(* IEC 61131-3 sources: 2026_Projet_YGO_ExcavatriceDragage/CODE_BACKUP/CODE_20260807_v0.5.25/COMMUN, 15 files *)

(* ---- E_State.st ---- *)
(* ═══════════════════════════════════════════════════════════════
   🚦 E_State — Phase opérationnelle d'un FB métier (valeurs EXCLUSIVES)
   ───────────────────────────────────────────────────────────────
    📄 Doc métier : DOC/AF_Partie-03_Contrats_Composants_v2.1.md §3
   ⚠️ Un seul état à la fois. Error / SafeStop / perte Enable sont
      ORTHOGONAUX à la phase (voir ErrorId, ne polluent pas State).
   🧩 Fondation manquante requise par le contrat FB (Partie3 §1).
   ═══════════════════════════════════════════════════════════════ *)

TYPE E_State :
ENUM
    DISABLED := 0,   (* Enable faux, neutralisé *)
    INIT     := 1,   (* Démarrage / vérifs *)
    READY    := 2,   (* Prêt, attend ordre *)
    BUSY     := 3,   (* Action en cours *)
    DONE     := 4,   (* Action terminée *)
    STOPPING := 5    (* Décél rampe avant arrêt (StartStop=FALSE ou SafeStop=TRUE) *)
END_ENUM
END_TYPE

(* ---- ST_ContactorCheck.st ---- *)
(* ═══════════════════════════════════════════════════════════════
   🔌 ST_ContactorCheck — Double vérification commande/retour contacteur
   ───────────────────────────────────────────────────────────────
    📄 Doc métier : DOC/AF_Partie-02_Architecture_Programme_v3.1.md §3,
                    DOC/AF_Partie-03_Contrats_Composants_v2.1.md §2
   Utilisé par FB_Brake (frein) et FB_Winch (contacteurs de sens) pour
   détecter un collage / une absence de fermeture d'un contacteur de
   puissance, au-delà d'un délai de cohérence (FeedbackTimeout du FB
   appelant).
   ═══════════════════════════════════════════════════════════════ *)

TYPE ST_ContactorCheck :
STRUCT
    Command     : BOOL;   // Ordre envoyé au contacteur (TRUE = fermé/actif)
    Feedback    : BOOL;   // Retour d'état câblé (TRUE = effectivement fermé)
    StuckClosed : BOOL;   // Diag : commande OFF mais retour ON depuis trop longtemps → PowerCutOff
    StuckOpen   : BOOL;   // Diag : commande ON mais retour OFF depuis trop longtemps
END_STRUCT
END_TYPE

(* ---- FB_Acquisition_Preflight.st ---- *)
(* ═══════════════════════════════════════════════════════════════
   🩺 FB_Acquisition_Preflight — Verdict passif machine arrêtée
   📄 Doc : ARCHIVES/Doc/AUDITS/PreLivraison/TASKS/TASK_D1_Preflight_et_Symetrie_Winch_v1.0.md
   🔒 Observateur pur : aucun SafeStop, PowerCutOff ou ordre machine.
   ═══════════════════════════════════════════════════════════════ *)
FUNCTION_BLOCK FB_Acquisition_Preflight
VAR_INPUT
    Execute : BOOL;
    MachineIsStill : BOOL;
    M1BrakeApplied, M2BrakeApplied, M3BrakeApplied : BOOL;
    M1ContactorsReleased, M2ContactorsReleased, M1ThermalOk, M2ThermalOk : BOOL;
    BrakeThermalOk, PhaseRotationOk, SlackCableTensioned, M3SensorWordIncoherent : BOOL;
    EmergencyChainClosed, PowerContactorEngaged, EncoderM1Operational, EncoderM2Operational : BOOL;
    HomedM1, HomedM2, M1PositionInBounds, M2PositionInBounds : BOOL;
END_VAR
VAR_OUTPUT
    PreflightOk : BOOL;
    PreflightDone : BOOL;
    PreflightBusy : BOOL;
    PreflightErrorId : WORD;
END_VAR
VAR
    ExecuteEdge : R_TRIG;
    BootPending : BOOL := TRUE;
    RequestPending : BOOL;
END_VAR

ExecuteEdge(CLK := Execute);
RequestPending := RequestPending OR ExecuteEdge.Q OR BootPending;
PreflightBusy := RequestPending AND NOT MachineIsStill;
IF NOT MachineIsStill THEN PreflightDone := FALSE; RETURN; END_IF;
IF NOT RequestPending THEN RETURN; END_IF;

PreflightErrorId := 0;
(* bit0..2 frein M1/M2/M3 serré; bit3..4 contacteurs M1/M2 retombés;
   bit5..6 thermique M1/M2 OK; bit7 thermique frein OK; bit8 phases OK;
   bit9 câble M2 tendu; bit10 mot M3 cohérent; bit11 contacteur sans chaîne;
   bit12..13 codeur M1/M2 opérationnel; bit14..15 homé et position bornée M1/M2. *)
IF NOT M1BrakeApplied THEN PreflightErrorId := PreflightErrorId OR 16#0001; END_IF;
IF NOT M2BrakeApplied THEN PreflightErrorId := PreflightErrorId OR 16#0002; END_IF;
IF NOT M3BrakeApplied THEN PreflightErrorId := PreflightErrorId OR 16#0004; END_IF;
IF NOT M1ContactorsReleased THEN PreflightErrorId := PreflightErrorId OR 16#0008; END_IF;
IF NOT M2ContactorsReleased THEN PreflightErrorId := PreflightErrorId OR 16#0010; END_IF;
IF NOT M1ThermalOk THEN PreflightErrorId := PreflightErrorId OR 16#0020; END_IF;
IF NOT M2ThermalOk THEN PreflightErrorId := PreflightErrorId OR 16#0040; END_IF;
IF NOT BrakeThermalOk THEN PreflightErrorId := PreflightErrorId OR 16#0080; END_IF;
IF NOT PhaseRotationOk THEN PreflightErrorId := PreflightErrorId OR 16#0100; END_IF;
IF NOT SlackCableTensioned THEN PreflightErrorId := PreflightErrorId OR 16#0200; END_IF;
IF M3SensorWordIncoherent THEN PreflightErrorId := PreflightErrorId OR 16#0400; END_IF;
IF PowerContactorEngaged AND NOT EmergencyChainClosed THEN PreflightErrorId := PreflightErrorId OR 16#0800; END_IF;
IF NOT EncoderM1Operational THEN PreflightErrorId := PreflightErrorId OR 16#1000; END_IF;
IF NOT EncoderM2Operational THEN PreflightErrorId := PreflightErrorId OR 16#2000; END_IF;
IF NOT HomedM1 OR NOT M1PositionInBounds THEN PreflightErrorId := PreflightErrorId OR 16#4000; END_IF;
IF NOT HomedM2 OR NOT M2PositionInBounds THEN PreflightErrorId := PreflightErrorId OR 16#8000; END_IF;
PreflightOk := (PreflightErrorId = 0); PreflightDone := TRUE; BootPending := FALSE; RequestPending := FALSE;

(* ---- FB_Brake.st ---- *)
(* ═══════════════════════════════════════════════════════════════
   🛑 FB_Brake — Séquence frein à manque de courant (temps physiques)
   ───────────────────────────────────────────────────────────────
   📄 Doc métier : DOC/AF_Partie-10_Fonction_Winch_v2.0.md §3
                   (règles issues de DOC/AF_Partie-04_Mode_SemiAuto_Sequenceur_v2.0.md §4)
   🛠️ Frein à manque de courant : colle au repos (sécurité positive).
   📥 MovementRequested : mouvement demandé par FB_Winch (sens+palier > 0)
   📤 BrakeCmd          : commande bobine frein — TRUE = relâché (alimenté)
   ⏱️ Séquence démarrage : attend fermeture contacteur + magnétisation
      moteur AVANT de relâcher (sinon charge retombe → à-coup).
   ⏱️ Séquence arrêt     : attend décélération/ouverture contacteur AVANT
      de coller (sinon usure/casse mécanique en plein mouvement).
   🔍 Double vérification retour contacteur bobine (ST_ContactorCheck) :
      incohérence commande/retour au-delà de FeedbackTimeout → ErrorId.
   🆕 REX 2026-08-03 (révocation 2026-07-26) : le retour câblé est l'image du CONTACTEUR DE COMMANDE
      (DI = 1 ⟺ frein ouvert). Plus d'inversion à la frontière : ce FB reçoit maintenant un
      signal dans le MÊME sens que `BrakeCmd` en marche saine (TRUE = relâché = ouvert) → le test d'incohérence est `<>`, pas `=`.
      ⚠️ Ce retour n'est PAS une mesure du frein : il détecte un contacteur/bobine défaillant, mais
      pas un frein usé ou qui patine. Le patinage reste couvert par Méca A (dérive codeur,
      FB_Safety_Winch bit7) — pas par ce bloc.
   ═══════════════════════════════════════════════════════════════ *)

// === DECLARATION (à coller dans la partie déclaration du POU FB_Brake) ===

FUNCTION_BLOCK PUBLIC FB_Brake
VAR_INPUT
    Enable              : BOOL;                     // Contexte général (comme tout FB) — FALSE = frein collé (sûr)
    Reset               : BOOL;                     // Acquittement défaut (front)
    MovementRequested   : BOOL;                      // TRUE = FB_Winch demande un mouvement (sens+palier actifs)
    ContactorFeedback   : BOOL;                      // Retour frein (`PRG_02_Acquisition.HwIn`) : TRUE = frein OUVERT (desserré)
                                                       // 🆕 REX 2026-08-03 : même sens que BrakeCmd (TRUE = relâché)
                                                       // → en marche normale les deux sont ÉGAUX ; c'est leur
                                                       //   DIFFÉRENCE qui trahit un contacteur collé (voir §4).
    DelayContactClose   : TIME := T#100ms;            // Temps de fermeture contacteur de puissance
    DelayMagnetise      : TIME := T#300ms;            // Délai magnétisation moteur avant ouverture frein
    DelayMotorDecel     : TIME := T#500ms;            // Délai décélération/ouverture contacteur avant collage frein
    FeedbackTimeout     : TIME := T#1s;               // Délai max cohérence commande/retour frein
    BypassContactorCheck: BOOL;                       // 🧪 TRUE = désactive StuckClosed/StuckOpen (axe simulé,
                                                       // voir GVL_Simulation.SensorMxContactorFeedbackIsReal, passé
                                                       // par l'appelant FB_Winch/FB_Translation — TOUJOURS FALSE réel)
END_VAR
VAR_OUTPUT
    Ready               : BOOL;
    Busy                : BOOL;
    Done                : BOOL;
    Error               : BOOL;
    ErrorId             : WORD;          // bit0: "Défaut engagement frein" - incohérence commande/retour frein (collage ou non-relâche)
    State               : E_State;
    StateAtError        : E_State;
    BrakeCmd            : BOOL;          // Commande sortie bobine frein : TRUE = relâché
    BrakeCommandOpenConfirmed : BOOL;    // TRUE = frein ouvert = commande ouverture confirmée (même sens que ContactorFeedback)
    ContactorCheck      : ST_ContactorCheck;  // Diag détaillé (IHM / FB_Safety_Winch)
END_VAR
VAR
    ResetEdge           : R_TRIG;
    ErrorEdge           : R_TRIG;
    BypassEdge          : R_TRIG;        // 🔑 REX 2026-07-24 : Front montant activation bypass pour réarmement immédiat
    TonMagnetise        : TON;           // Temporisation avant relâche
    TonDecel            : TON;           // Temporisation avant collage
    TonFeedback         : TON;           // Timeout cohérence commande/retour
END_VAR

// === IMPLEMENTATION (à coller dans le corps ST du POU FB_Brake) ===

// 🛑 1. GATE — pas d'Enable = frein collé (sécurité positive), aucune temporisation en cours
IF NOT Enable THEN
    TonMagnetise(IN := FALSE, PT := DelayMagnetise + DelayContactClose);
    TonDecel(IN := FALSE, PT := DelayMotorDecel);
    BrakeCmd := FALSE;
    State := E_State.DISABLED;
    Ready := FALSE; Busy := FALSE; Done := FALSE;
    RETURN;
END_IF;

Ready := TRUE;

// 🔑 2. RESET FRONT — efface le bit dont la cause a disparu
ResetEdge(CLK := Reset);
BypassEdge(CLK := BypassContactorCheck);

// 🛠️ 3. SÉQUENCE TEMPORISÉE (démarrage vs arrêt)
IF MovementRequested THEN
    TonDecel(IN := FALSE, PT := DelayMotorDecel);
    TonMagnetise(IN := TRUE, PT := DelayMagnetise + DelayContactClose);
    IF TonMagnetise.Q THEN
        BrakeCmd := TRUE;              // ✅ Contacteur + magnétisation acquis → relâche
        State := E_State.DONE;
    ELSE
        BrakeCmd := FALSE;             // ⏳ Encore collé pendant la magnétisation
        State := E_State.BUSY;
    END_IF;
ELSE
    // 🆕 REX 2026-07-08 : Sécurité positive - fermeture immédiate du frein (collé) dès que les contacteurs de sens s'ouvrent
    TonMagnetise(IN := FALSE, PT := DelayMagnetise + DelayContactClose);
    TonDecel(IN := FALSE, PT := DelayMotorDecel);
    BrakeCmd := FALSE;                 // Fermeture immédiate
    State := E_State.READY;
END_IF;

Busy := (State = E_State.BUSY);
Done := (State = E_State.DONE);

// 🔍 4. DOUBLE VÉRIFICATION RETOUR CONTACTEUR (ST_ContactorCheck)
ContactorCheck.Command := BrakeCmd;
ContactorCheck.Feedback := ContactorFeedback;

// 🆕 REX 2026-08-03 (révocation 2026-07-26) : `ContactorFeedback` est maintenant dans le MÊME sens
// que `BrakeCmd` (TRUE = relâché = frein ouvert). En marche saine les deux sont ÉGAUX → c'est leur
// DIFFÉRENCE qui signale l'incohérence (contacteur collé).
// ⚠️ Le test repasse en `<>` (retour à la logique d'origine pré-2026-07-26).
TonFeedback(IN := (BrakeCmd <> ContactorFeedback), PT := FeedbackTimeout);
IF NOT BypassContactorCheck THEN
    IF TonFeedback.Q THEN
        ContactorCheck.StuckClosed := (BrakeCmd AND NOT ContactorFeedback);            // relâche commandée (BrakeCmd=TRUE), frein reste serré (ContactorFeedback=FALSE)
        ContactorCheck.StuckOpen   := (NOT BrakeCmd AND ContactorFeedback);             // serrage commandé (BrakeCmd=FALSE), frein reste ouvert (ContactorFeedback=TRUE)
        ErrorId := ErrorId OR 16#0001;
    ELSIF ResetEdge.Q THEN
        ContactorCheck.StuckClosed := FALSE;
        ContactorCheck.StuckOpen   := FALSE;
        ErrorId := ErrorId AND 16#FFFE;
    END_IF;
ELSE
    ContactorCheck.StuckClosed := FALSE;
    ContactorCheck.StuckOpen   := FALSE;
    ErrorId := ErrorId AND 16#FFFE;   // Bypass actif : efface/maintient à 0 le bit 0
    IF BypassEdge.Q THEN
        StateAtError := E_State.DISABLED; // Front activation bypass : débloque l'état figé
    END_IF;
END_IF;

// 🧾 5. ARBITRAGE ERROR / STATEATERROR (figé jusqu'à acquittement)
Error := (ErrorId <> 16#0000);
ErrorEdge(CLK := Error);
IF ErrorEdge.Q THEN
    StateAtError := State;
END_IF;

// 🛡️ 6. SORTIE SÛRE SUR DÉFAUT
IF Error THEN
    BrakeCmd := FALSE;
END_IF;

// 📤 7. CONFIRMATION OUVERTURE FREIN (même sens que ContactorFeedback, ou image de BrakeCmd si BypassContactorCheck=TRUE)
IF BypassContactorCheck THEN
    BrakeCommandOpenConfirmed := BrakeCmd;
ELSE
    BrakeCommandOpenConfirmed := ContactorFeedback;  (* TRUE = frein ouvert = desserrage confirmé *)
END_IF;

(* ---- FB_CfgPersistBridge_BucketCfg.st ---- *)
(* ═══════════════════════════════════════════════════════════════
   🌉 FB_CfgPersistBridge_BucketCfg — Pont persistance générique pour ST_BucketCfg
   ───────────────────────────────────────────────────────────────
   🎯 Voir FB_CfgPersistBridge_SyncCfg.st (Lot 3a) pour la logique de référence — identique,
   seul le type ST_BucketCfg change. La copie struct-à-struct gère aussi le sous-struct imbriqué
   Config : ST_BucketConfig automatiquement (pas de traitement spécial nécessaire).
   ═══════════════════════════════════════════════════════════════ *)
FUNCTION_BLOCK FB_CfgPersistBridge_BucketCfg
VAR_IN_OUT
    Hmi     : ST_BucketCfg; (* 🖥️ ex. GVL_IHM.M2TreuilBenne.Bucket.Cfg *)
    Persist : ST_BucketCfg; (* 💾 ex. GVL_PERSISTENT._BucketCfgPersist *)
END_VAR
VAR_OUTPUT
    JustRestored : BOOL;
END_VAR

JustRestored := FALSE;
IF NOT Hmi.Initialized THEN
    Hmi := Persist;
    Hmi.Initialized := TRUE;
    JustRestored := TRUE;
ELSE
    Persist := Hmi;
END_IF;

(* ---- FB_CfgPersistBridge_CommunCfg.st ---- *)
(* ═══════════════════════════════════════════════════════════════
   🌉 FB_CfgPersistBridge_CommunCfg — Pont persistance générique pour ST_CommunCfg
   ───────────────────────────────────────────────────────────────
   🎯 Voir FB_CfgPersistBridge_SyncCfg.st (Lot 3a) pour la logique de référence — identique,
   seul le type ST_CommunCfg change.
   ═══════════════════════════════════════════════════════════════ *)
FUNCTION_BLOCK FB_CfgPersistBridge_CommunCfg
VAR_IN_OUT
    Hmi     : ST_CommunCfg; (* 🖥️ ex. GVL_IHM.Commun.Cfg *)
    Persist : ST_CommunCfg; (* 💾 ex. GVL_PERSISTENT._CommunCfgPersist *)
END_VAR
VAR_OUTPUT
    JustRestored : BOOL;
END_VAR

JustRestored := FALSE;
IF NOT Hmi.Initialized THEN
    Hmi := Persist;
    Hmi.Initialized := TRUE;
    JustRestored := TRUE;
ELSE
    Persist := Hmi;
END_IF;

(* ---- FB_CfgPersistBridge_CycleCfg.st ---- *)
(* ═══════════════════════════════════════════════════════════════
   🌉 FB_CfgPersistBridge_CycleCfg — Pont persistance générique pour ST_CycleCfg
   ───────────────────────────────────────────────────────────────
   🎯 Voir FB_CfgPersistBridge_SyncCfg.st (Lot 3a) pour la logique de référence — identique,
   seul le type ST_CycleCfg change.
   ═══════════════════════════════════════════════════════════════ *)
FUNCTION_BLOCK FB_CfgPersistBridge_CycleCfg
VAR_IN_OUT
    Hmi     : ST_CycleCfg; (* 🖥️ ex. GVL_IHM.Cycle.Cfg *)
    Persist : ST_CycleCfg; (* 💾 ex. GVL_PERSISTENT._CycleCfgPersist *)
END_VAR
VAR_OUTPUT
    JustRestored : BOOL;
END_VAR

JustRestored := FALSE;
IF NOT Hmi.Initialized THEN
    Hmi := Persist;
    Hmi.Initialized := TRUE;
    JustRestored := TRUE;
ELSE
    Persist := Hmi;
END_IF;

(* ---- FB_CfgPersistBridge_DredgingAssistCfg.st ---- *)
(* ═══════════════════════════════════════════════════════════════
   🌉 FB_CfgPersistBridge_DredgingAssistCfg — Pont IHM/persistance prélèvement
   ═══════════════════════════════════════════════════════════════ *)
FUNCTION_BLOCK FB_CfgPersistBridge_DredgingAssistCfg
VAR_IN_OUT
    Hmi     : ST_DredgingAssistCfg;
    Persist : ST_DredgingAssistCfg;
END_VAR
VAR_OUTPUT
    JustRestored : BOOL;
END_VAR

JustRestored := FALSE;
IF NOT Hmi.Initialized THEN
    Hmi := Persist;
    Hmi.Initialized := TRUE;
    JustRestored := TRUE;
ELSE
    Persist := Hmi;
END_IF;

(* ---- FB_CfgPersistBridge_SyncCfg.st ---- *)
(* ═══════════════════════════════════════════════════════════════
   🌉 FB_CfgPersistBridge_SyncCfg — Pont persistance générique pour ST_SyncCfg
   ───────────────────────────────────────────────────────────────
   🎯 Remplace les blocs manuels restauration/sauvegarde dupliqués à chaque domaine
   (voir DOC/AUDITS/ConfigPersistence/). Une instance = un couple (struct IHM, struct
   GVL_PERSISTENT) du MÊME type. Logique :
   - Hmi.Initialized = FALSE (RETAIN invalidé, ex. changement de layout DUT) → restaure
     Hmi depuis Persist, marque Initialized, pulse JustRestored 1 scan.
   - Hmi.Initialized = TRUE → sauvegarde continue Hmi vers Persist (jamais l'inverse).
   🔒 Défense en profondeur : jamais d'écriture PERSISTENT avant qu'une restauration
   réussie n'ait eu lieu (même principe que tous les blocs Cfg du Lot 2).
   ═══════════════════════════════════════════════════════════════ *)
FUNCTION_BLOCK FB_CfgPersistBridge_SyncCfg
VAR_IN_OUT
    Hmi     : ST_SyncCfg; (* 🖥️ ex. GVL_IHM.M1M2Sync.Cfg — struct exposé à l'IHM *)
    Persist : ST_SyncCfg; (* 💾 ex. GVL_PERSISTENT._SyncCfgPersist — mémoire PERSISTENT *)
END_VAR
VAR_OUTPUT
    JustRestored : BOOL; (* 🔔 TRUE pendant 1 scan le boot où la restauration a eu lieu —
                             l'appelant s'en sert pour piloter GVL_IHM.Commun.ConfigRestoredFromPersistent *)
END_VAR

JustRestored := FALSE;
IF NOT Hmi.Initialized THEN
    Hmi := Persist;
    Hmi.Initialized := TRUE;
    JustRestored := TRUE;
ELSE
    Persist := Hmi;
END_IF;

(* ---- FB_CfgPersistBridge_TranslationCfg.st ---- *)
(* ═══════════════════════════════════════════════════════════════
   🌉 FB_CfgPersistBridge_TranslationCfg — Pont persistance générique pour ST_TranslationCfg
   ───────────────────────────────────────────────────────────────
   🎯 Instance unique : TranslationM3.Cfg (un seul axe M3, contrairement à M1/M2).
   Restaure Persist → Hmi au boot si nécessaire, puis sauvegarde Hmi → Persist.
   ═══════════════════════════════════════════════════════════════ *)
FUNCTION_BLOCK FB_CfgPersistBridge_TranslationCfg
VAR_IN_OUT
    Hmi     : ST_TranslationCfg; (* 🖥️ Struct exposé à l'IHM *)
    Persist : ST_TranslationCfg; (* 💾 Mémoire PERSISTENT *)
END_VAR
VAR_OUTPUT
    JustRestored : BOOL; (* 🔔 TRUE pendant le scan de restauration *)
END_VAR

JustRestored := FALSE;
IF NOT Hmi.Initialized THEN
    Hmi := Persist;
    Hmi.Initialized := TRUE;
    JustRestored := TRUE;
ELSE
    Persist := Hmi;
END_IF;

(* ---- FB_CfgPersistBridge_WinchCfg.st ---- *)
(* ═══════════════════════════════════════════════════════════════
   🌉 FB_CfgPersistBridge_WinchCfg — Pont persistance générique pour ST_WinchCfg
   ───────────────────────────────────────────────────────────────
   🎯 Deux instances indépendantes : M1TreuilRetenue.Cfg et M2TreuilBenne.Cfg.
   Restaure Persist → Hmi au boot si nécessaire, puis sauvegarde Hmi → Persist.
   ═══════════════════════════════════════════════════════════════ *)
FUNCTION_BLOCK FB_CfgPersistBridge_WinchCfg
VAR_IN_OUT
    Hmi     : ST_WinchCfg; (* 🖥️ Struct exposé à l'IHM *)
    Persist : ST_WinchCfg; (* 💾 Mémoire PERSISTENT *)
END_VAR
VAR_OUTPUT
    JustRestored : BOOL; (* 🔔 TRUE pendant le scan de restauration *)
END_VAR

JustRestored := FALSE;
IF NOT Hmi.Initialized THEN
    Hmi := Persist;
    Hmi.Initialized := TRUE;
    JustRestored := TRUE;
ELSE
    Persist := Hmi;
END_IF;

(* ---- FB_CycleTime.st ---- *)
(* ═══════════════════════════════════════════════════════════════
   ⏱️ FB_CycleTime — Mesure du temps de cycle réel de la tâche
   ───────────────────────────────────────────────────────────────
   📄 Doc métier : DOC/AF_Partie-08_Fonction_Joystick_v2.0.md §2
      (base de temps utilisée par FB_Filter_PT1, composé dans FB_Joystick)
   ═══════════════════════════════════════════════════════════════ *)
FUNCTION_BLOCK FB_CycleTime
VAR_INPUT
    DefaultValueS : REAL := 0.004; (* Valeur de secours par défaut (ex. 4ms) *)
END_VAR
VAR_OUTPUT
    CycleTimeS    : REAL;          (* Temps écoulé réel calculé (secondes) *)
END_VAR
VAR
    TimeCurrent   : TIME;          (* Temps système actuel *)
    TimeLast      : TIME;          (* Empreinte de temps du cycle précédent *)
    DeltaTimeMs   : UDINT;         (* Écart brut calculé (ms) *)
    InitDone      : BOOL;          (* Drapeau d'initialisation du premier cycle *)
END_VAR

// 1. ACQUISITION DU TEMPS SYSTÈME
TimeCurrent := TIME();

// 2. INITIALISATION UNIQUE AU PREMIER CYCLE
IF NOT InitDone THEN
    TimeLast := TimeCurrent;
    InitDone := TRUE;
    CycleTimeS := DefaultValueS;
    RETURN;
END_IF;

// 3. CALCUL DU DELTA EN MILLISECONDES
DeltaTimeMs := TIME_TO_UDINT(TimeCurrent - TimeLast);

// 4. CONVERSION ET CHARGE DE SECOURS
IF DeltaTimeMs > 0 THEN
    CycleTimeS := UDINT_TO_REAL(DeltaTimeMs) / 1000.0;
ELSE
    CycleTimeS := DefaultValueS;
END_IF;

// 5. ARCHIVAGE POUR LE PROCHAIN CYCLE
TimeLast := TimeCurrent;

(* ---- FB_DigitalInputFilter.st ---- *)
(* ═══════════════════════════════════════════════════════════════
   📥 FB_DigitalInputFilter — Filtre temporel minimal d'une entrée TOR
   ───────────────────────────────────────────────────────────────
   📄 Doc : DOC/AF_Partie-06_Acquisition_Qualification_IO_v2.1.md
   🎯 Rôle unique : accepter un changement BOOL seulement après FilterTime.
   🛡️ Ce FB ne normalise pas la polarité et ne réalise aucun diagnostic device.
      La polarité est portée par le nom/mapping d'acquisition ; la santé carte
      est publiée séparément par PRG_02_Acquisition.GetDeviceState().
   🔗 Producteur : PRG_02_Acquisition, image HwRealQualified.
   ═══════════════════════════════════════════════════════════════ *)

FUNCTION_BLOCK PUBLIC FB_DigitalInputFilter
VAR_INPUT
    InputRaw   : BOOL; (* Valeur brute du canal réel *)
    FilterTime : TIME; (* Durée minimale de stabilité avant validation *)
END_VAR
VAR_OUTPUT
    State : BOOL; (* Valeur filtrée ; première valeur prise immédiatement au démarrage *)
END_VAR
VAR
    FilterTon     : TON;
    FirstScanDone : BOOL;
END_VAR

IF NOT FirstScanDone THEN
    State := InputRaw;
    FirstScanDone := TRUE;
ELSE
    FilterTon(IN := (InputRaw <> State), PT := FilterTime);
    IF FilterTon.Q THEN
        State := InputRaw;
    END_IF;
END_IF;

(* ---- FB_Output.st ---- *)
(* ═══════════════════════════════════════════════════════════════
   📤 FB_Output — Sortie relais (brique réduite, REX 2026-08-04)
   ───────────────────────────────────────────────────────────────
   📄 Doc métier : DOC/AF_Partie-03_Contrats_Composants_v2.1.md §Câblage
   🧭 Interface RÉDUITE (validée utilisateur 2026-08-04) : relais de
      commande BAS NIVEAU — transmet fidèlement `Command` (déjà
      résolu/rampé par le FB métier appelant), ne décide JAMAIS lui-même
      d'un arrêt de mouvement.
   🔁 Rôle : inversion NO/NC uniquement.
   🗑️ REX 2026-08-04 : partie FEEDBACK retirée (FeedbackRaw, UseFeedback,
      Blink1Hz, FeedbackTimeout, ChannelOk, FeedbackOk, Error, ErrorId) —
      jamais câblée (0 usage dans PRG_06, 15 instances Command→State).
      Diagnostic contacteur déjà couvert au niveau métier par
      FB_Safety_Winch (FwdRevSpeedFeedbackOff, BrakeFeedback).
   ═══════════════════════════════════════════════════════════════ *)

FUNCTION_BLOCK PUBLIC FB_Output
VAR_INPUT
    Command     : BOOL;   // Ordre logique, déjà résolu/rampé par le FB métier appelant
    InvertLogic : BOOL;   // TRUE = câblage NC (inversion de la sortie)
END_VAR
VAR_OUTPUT
    State       : BOOL;   // Vers la carte de sortie
END_VAR

// === IMPLEMENTATION (à coller dans le corps ST du POU FB_Output) ===

State := Command XOR InvertLogic;

(* ---- FB_Ramp.st ---- *)
(* ═══════════════════════════════════════════════════════════════
   📈 FB_Ramp — Rampe accel/décel anti-à-coups (retour zéro plus rapide)
   ───────────────────────────────────────────────────────────────
   📄 Doc métier : DOC/AF_Partie-08_Fonction_Joystick_v2.0.md §2 (usage),
                   DOC/AF_Partie-10_Fonction_Winch_v2.0.md (correctif ci-dessous)
   🧩 Instancié 3 fois dans le projet : RampX/RampY (FB_Joystick, cible
      SIGNÉE -100..+100 %) et SpeedRamp (FB_Winch, cible TOUJOURS >= 0,
      jamais concernée par ce bug — voir analyse d'impact ci-dessous).

   ⚠️ CORRECTIF (retour terrain 2026-07-02) : le choix accel/décel
   comparait `Target`/`Current` AVEC LEUR SIGNE, pas leur magnitude.
   Conséquence : lors d'une inversion RAPIDE du joystick (Current très
   négatif, Target qui redevient positif), la condition
   `(Target > 0.0 AND Target > Current)` devenait vraie dès que `Target`
   passait légèrement positif — alors que `Current` était encore très
   loin de zéro côté négatif — et sélectionnait à tort `AccelRate` (lent,
   "s'éloigne du zéro") au lieu de `DecelRate` (rapide, "retourne vers le
   zéro") pour toute la portion du trajet qui ramène réellement vers
   zéro. Résultat observé : lors d'un flick rapide du joystick, `Current`
   mettait ~3× plus longtemps que prévu à repasser par zéro, ce qui
   retardait en cascade `AxisCmdY.Direction`/`SpeedRef`, puis l'interlock
   de sens de `FB_Winch` (`CommandedDirection` bloqué sur l'ancien sens
   plus longtemps que nécessaire).
   🔬 Analyse d'impact (avant correctif) : `FB_Ramp` n'est instancié que
   dans `FB_Joystick` (`RampX`/`RampY`, cible signée → CONCERNÉ) et dans
   `FB_Winch` (`SpeedRamp`, cible = `RampTargetPct` toujours >= 0 → JAMAIS
   de traversée de signe possible → NON concerné, comportement inchangé).
   ✅ Correction : classification basée sur le CÔTÉ de zéro où se trouve
   `Current` et le sens de déplacement (pas le signe brut de `Target`),
   vérifiée sur les 8 cas (Current>0/<0/=0 × s'éloigne/retourne/traverse).
   ═══════════════════════════════════════════════════════════════ *)

// === DECLARATION (à coller dans la partie déclaration du POU FB_Ramp) ===

FUNCTION_BLOCK FB_Ramp
VAR_INPUT
    Target      : REAL;       // Cible visée
    AccelRate   : REAL;       // Taux d'accélération (%/s)
    DecelRate   : REAL;       // Taux de décélération (%/s)
    CycleTimeS  : REAL;       // Temps de cycle réel en secondes
END_VAR
VAR_OUTPUT
    Current     : REAL;       // Valeur courante amortie
END_VAR
VAR
    StepX       : REAL;
    TargetLimited : REAL;
END_VAR

// === IMPLEMENTATION (à coller dans le corps ST du POU FB_Ramp) ===

// Détection du comportement (Accélération vs Décélération)
// 🔧 CORRECTIF : classification par CÔTÉ DE ZÉRO + sens de déplacement, plus par signe brut
// de Target seul (l'ancienne version se trompait lors d'une traversée de zéro rapide).
// 🛡️ Garde-fou : la rampe ne sort jamais de la plage normalisée ±100 %.
TargetLimited := LIMIT(-100.0, Target, 100.0);
Current := LIMIT(-100.0, Current, 100.0);

IF (Current >= 0.0 AND TargetLimited >= Current) OR (Current <= 0.0 AND TargetLimited <= Current) THEN
    StepX := AccelRate * CycleTimeS; // S'éloigne du zéro (reste du même côté, va plus loin)
ELSE
    StepX := DecelRate * CycleTimeS; // Retourne vers zéro, ou le traverse vers l'autre signe
END_IF;

// Application de la rampe
IF Current < TargetLimited THEN
    Current := Current + StepX;
    IF Current > TargetLimited THEN Current := TargetLimited; END_IF;
ELSIF Current > TargetLimited THEN
    Current := Current - StepX;
    IF Current < TargetLimited THEN Current := TargetLimited; END_IF;
END_IF;

// 🛡️ Limitation finale : même une valeur d'état déjà corrompue reste bornée.
Current := LIMIT(-100.0, Current, 100.0);
